Fanuc KAREL source: kt00416.KL

-- PROVISIONAL review KL for V770-1; original PC SHA256 2526e92b8b6dee1773b1a2e86352b53111622762f802385b67d8b4b8bca484ef
-- Incomplete behavior may be omitted. Consult companion uncertainty JSON. Do not deploy.
PROGRAM KT00416
%NOLOCKGROUP
VAR
  R2 : REAL
  OUT : BOOLEAN
-- UNRESOLVED_DECL H1 type=002017
BEGIN
  -- UNRESOLVED_PC offsets 5-19; opcodes 2E,22,9D,33,B4
  -- UNRESOLVED_PC offsets 24-35; opcodes 2E,23
  -- UNRESOLVED_PC offsets 40-65; opcodes 22,9D,33,B3,21,29,64,29,71,23
  -- UNRESOLVED_PC offsets 70-74; opcodes 7F
END KT00416
